(* IEC 61131-3 sources: plc-workbench/experiments/general_tasks_r6/final_recheck/interlocked_start, 2 files *)

(* ---- before.st ---- *)
FUNCTION_BLOCK InterlockedStart
VAR_INPUT
    start : BOOL;
    stop : BOOL;
    permit : BOOL;
END_VAR
VAR_OUTPUT
    running : BOOL;
END_VAR
VAR
    previousStart : BOOL := FALSE;
    startRising : BOOL;
END_VAR

startRising := start AND NOT previousStart;
previousStart := start;

IF stop OR NOT permit THEN
    running := FALSE;
ELSIF startRising THEN
    running := TRUE;
END_IF;

END_FUNCTION_BLOCK

(* ---- candidate_final.st ---- *)
FUNCTION_BLOCK InterlockedStart
VAR_INPUT
    start : BOOL;
    stop : BOOL;
    permit : BOOL;
END_VAR
VAR_OUTPUT
    running : BOOL;
END_VAR
VAR
    previousStart : BOOL := FALSE;
    startRising : BOOL;
END_VAR

startRising := start AND NOT previousStart;
previousStart := start;

IF stop OR NOT permit THEN
    running := FALSE;
ELSIF startRising THEN
    running := TRUE;
END_IF;

END_FUNCTION_BLOCK
